SUBAPPLICATION Uebung_OPC_L02_AX (* Wie Training_02 (Protokoll-FBs direkt statt im Composite), lokal: logiBUS_IXA -> AX_PUBLISH_1, AX_SUBSCRIBE_1 -> logiBUS_QXA *)
  (* Standard: 61499-2; Description: Copyright (c) 2026 Meisterschulen am Ostbahnhof This program and the accompanying materials are made available under the terms of the Eclipse Public License 2.0 which is available at https://www.eclipse.org/legal/epl-2.0/ SPDX-License-Identifier: EPL-2.0 *)
  (* Version 1.0, 2026-10-18, Franz Höpfinger, Meisterschulen am Ostbahnhof, OPC-UA lokal auf einem Geraet (Meins/OPC_UA_Lokal) *)
  PACKAGE Meins::OPC_UA_Lokal;
  IMPORT Meins::OPC_UA_Lokal::const::OpcUaLokal::Q1_WRITE;
  IMPORT Meins::OPC_UA_Lokal::const::OpcUaLokal::Q1_READ;
  IMPORT logiBUS::io::DI::logiBUS_DI::Input_I1;
  IMPORT logiBUS::io::DQ::logiBUS_DO::Output_Q1;
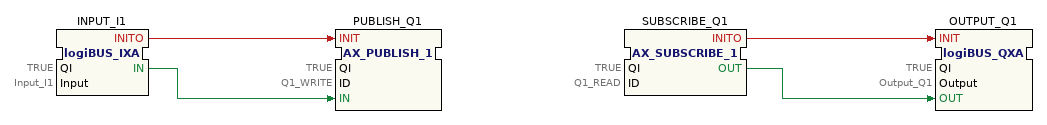
  FBS
    INPUT_I1 : logiBUS::io::DI::logiBUS_IXA(QI := TRUE, Input := Input_I1);
    PUBLISH_Q1 : adapter::net::AX_PUBLISH_1(QI := TRUE, ID := Q1_WRITE);
    SUBSCRIBE_Q1 : adapter::net::AX_SUBSCRIBE_1(QI := TRUE, ID := Q1_READ);
    OUTPUT_Q1 : logiBUS::io::DQ::logiBUS_QXA(QI := TRUE, Output := Output_Q1);
  END_FBS
  EVENT_CONNECTIONS
    INPUT_I1.INITO TO PUBLISH_Q1.INIT;
    SUBSCRIBE_Q1.INITO TO OUTPUT_Q1.INIT;
  END_CONNECTIONS
  ADAPTER_CONNECTIONS
    INPUT_I1.IN TO PUBLISH_Q1.IN;
    SUBSCRIBE_Q1.OUT TO OUTPUT_Q1.OUT;
  END_CONNECTIONS
END_SUBAPPLICATION
